(* IEC 61131-3 sources: trust-platform/examples/memory_marker_counter/src, 2 files *)

(* ---- Configuration.st ---- *)
CONFIGURATION MarkerCounter
TASK Cycle (INTERVAL := T#50ms, PRIORITY := 1);
PROGRAM P1 WITH Cycle : MainProgram;
VAR_CONFIG
    P1.Counter AT %MW0 : INT;
    P1.CounterLatched AT %QW0 : INT;
END_VAR
END_CONFIGURATION

(* ---- Main.st ---- *)
PROGRAM MainProgram
VAR
    Counter : INT;
    CounterLatched : INT;
END_VAR

CounterLatched := Counter;
Counter := Counter + 1;
END_PROGRAM
